{region 'Documentation'}
(*!
<summary>Check that IN is greater than Minimum.</summary>
*)
{endregion}
FUNCTION_BLOCK AssertGreaterThan_LInt EXTENDS AssertionBase
VAR_INPUT
    IN : LINT; //! Actual value checked or observed by this Assertion.
    Minimum : LINT; //! Exclusive lower bound; the actual value or count must be greater.
END_VAR

SUPER^();

{region 'Documentation'}
(*!
<summary>Check that IN is greater than Minimum.</summary>
*)
{endregion}
METHOD PROTECTED Assert
VAR
    Message : STRING(GVL_Constants.MessageLength);
    MinimumText : STRING(GVL_Constants.AssertionValueLength);
    ActualText : STRING(GVL_Constants.AssertionValueLength);
END_VAR
IF NOT EvaluationActive THEN
    RETURN;
END_IF;

IF Result = E_Result.Error THEN
    RETURN;
END_IF;

IF Result = E_Result.Failed THEN
    RETURN;
END_IF;

IF IN <= Minimum THEN
    MinimumText := LINT_TO_STRING(Minimum);
    ActualText := LINT_TO_STRING(IN);
    Message := CONCAT('Assertion failed: value is not greater than minimum. Minimum = ',
        MinimumText);
    Message := CONCAT(Message, ', Actual = ');
    Message := CONCAT(Message, ActualText);
    Message := CONCAT(Message, '.');
    Fail(Message := Message);
    RETURN;
END_IF;

Pass();
END_METHOD

END_FUNCTION_BLOCK

(* stored: Version 1.1.0.1
   POU AssertGreaterThan_LInt: Id {91c17091-ac5e-4b1c-b7e8-3ac0f801b2e1}, SpecialFunc None
   Folder Internal: Id {affcc26e-dbab-4718-9c4f-7ef421a93f9c}
   Method Assert: Id {8cd8a8b9-6946-453b-972a-8155fc787ebc} *)
